// Mitsubishi GX Works2 project: 261019_특수기능타이머(STMR)   PLC: Q03UDV

PROGRAM MAIN
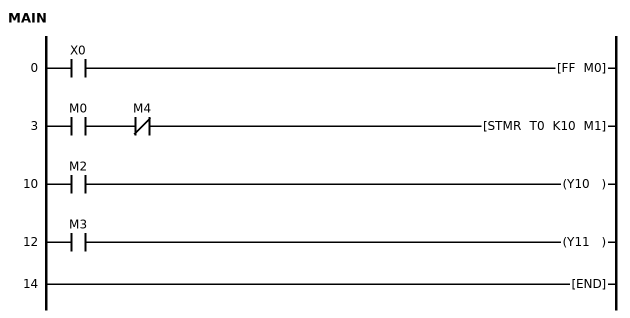
0     LD      X0
      FF      M0
3     LD      M0
      ANI     M4
      STMR    T0 K10 M1
10    LD      M2
      OUT     Y10
12    LD      M3
      OUT     Y11
14    END
END_PROGRAM
